{attribute 'qualified_only'}
VAR_GLOBAL CONSTANT
    startDelay : TIME := T#1s;
END_VAR

(* stored: Version 1.1.0.1, ProductVersion 3.1 *)
